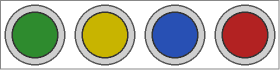
VISUALIZATION vis_Cycle_Panel  // 280x70
VAR_IN_OUT
	fb: FB_SFC_Cycle;
END_VAR
    Lamp1 (0,0 70x70), tooltip "Ready", variable: fb.bReady, style: Lamp-Lamp1-Green
    Lamp1 (70,0 70x70), tooltip "Done", variable: fb.bDone, style: Lamp-Lamp1-Yellow
    Lamp1 (140,0 70x70), tooltip "ToBe Done", variable: fb.bToBe_Done, style: Lamp-Lamp1-Blue
    Lamp1 (210,0 70x70), tooltip "Run", variable: fb.bRun, style: Lamp-Lamp1-Red
END_VISUALIZATION

(* stored: Version 1.1.0.1, ProductVersion 3.1.4024.12
   Visu vis_Cycle_Panel: Id {6b7e133d-15a5-4167-b20f-033efbef6c2b} *)
